// TwinCAT 3 PLC project Untitled1
// ProgramVersion: 3.1.4026.26
// project tree:
//   GVLs/HMI/ CNV_HMI.TcGVL, CNV_HMI_IO.TcGVL, GVL_HMI_Carousel.TcGVL, GVL_HMI_CNV.TcGVL, GVL_HMI_Gates.TcGVL, GVL_HMI_System.TcGVL, GVL_HMI_VTD.TcGVL
//   GVLs/IO/ IO_Cards.TcGVL, IO_Chargers.TcGVL, IO_RemoteModules.TcGVL, IO_Safety.TcGVL, IO_VFDs.TcGVL

// ---- GVLs/HMI/CNV_HMI.TcGVL
{attribute 'qualified_only'}
VAR_GLOBAL
	CNV_ID_HMI_Old_1:  DINT;
	CNV_ID_HMI:  DINT;
	CNV_ID_HMI_1:  DINT;
	CNV_ID_HMI_Old:  DInt;
	CNV_In_Out_1:  BOOL;
	CNV_Level_Selected:  UInt;
	CNV_Level_Selected_OLD:  UInt;
	CNV_Motor_Actual_Torque:  Real;
	CNV_Motor_Actual_Torque_1:  REAL;
	CNV_Motor_Current_Actual_HMI:  Real;
	CNV_Motor_Current_Actual_HMI_1:  REAL;
	CNV_Motor_Ready:  Bool;
	CNV_Motor_Ready_1:  BOOL;
	CNV_Motor_Status_HMI:  UInt;
	CNV_Motor_Status_HMI_1:  UINT;
	Cnv_Occupied_HMI:  Bool;
	Cnv_Occupied_HMI_1:  BOOL;
	CNV_System_Selected:  UInt;
	CVTD_CNV2_Selected:  UInt;
	Enable_HMI:  Bool;
	Enable_HMI_1:  Bool;
	Enabled_HMI:  Bool;
	Enabled_HMI_1:  Bool;
	Error_HMI:  Bool;
	Error_HMI_1:  Bool;
	HMI_Light_Guard_Bypass:  Bool;
	Light_Guard_Bypass_1:  Bool;
	Light_Guard_Bypass_2:  Bool;
	Manual_Bwd_HMI:  Bool;
	Manual_Bwd_HMI_1:  Bool;
	Manual_Fwd_HMI:  Bool;
	Manual_Fwd_HMI_1:  Bool;
	Manual_Sfty_Stopper_Down_1:  Bool;
	Manual_Sfty_Stopper_Up_1:  Bool;
	Mode_Change_HMI:  UInt;
	Mode_Change_HMI_1:  UInt;
	Mode_HMI:  UInt;
	Mode_HMI_1:  UInt;
	Motor_Direction_HMI:  UInt;
	Motor_Direction_HMI_1:  UInt;
	Motor_Speed_Actual_HMI:  UInt;
	Motor_Speed_Actual_HMI_1:  UInt;
	Motor_Speed_Requested_HMI:  UInt;
	Motor_Speed_Requested_HMI_1:  UInt;
	Ready_For_Task_HMI:  Bool;
	Ready_For_Task_HMI_1:  Bool;
	Reset_HMI:  Bool;
	Reset_HMI_1:  Bool;
	Running_HMI:  Bool;
	Running_HMI_1:  Bool;
	SM_State_HMI:  UInt;
	SM_State_HMI_1:  UInt;
	Start_Transfer_HMI:  Bool;
	Start_Transfer_HMI_1:  Bool;
	Stop_HMI:  Bool;
	Stopped_HMI:  Bool;
	Stopped_HMI_1:  Bool;
	Transfer_From_ID_HMI:  DInt;
	Transfer_From_ID_HMI_1:  DInt;
	Transfer_To_ID_HMI:  DInt;
	Transfer_To_ID_HMI_1:  DInt;
	UpDown_1:  UInt;
	Warning_HMI:  UInt;
	Warning_HMI_1:  UINT;
END_VAR

// ---- GVLs/HMI/CNV_HMI_IO.TcGVL
{attribute 'qualified_only'}
VAR_GLOBAL
	HMI_CNV_SftyPinDown_1:  BOOL;
	HMI_CNV_SftyPinUp_1:  BOOL;
	HMI_Light_Guard:  Bool;
	HMI_CNV_Forward_1:  Bool;
	HMI_CNV_Backward:  Bool;
	HMI_CNV_Forward:  Bool;
	HMI_CNV_Backward_1:  Bool;
END_VAR

// ---- GVLs/HMI/GVL_HMI_Carousel.TcGVL
// HMI interface of the screen Carrousel.
// Device index: 1..2 = PopUp 1..2, 3..7 = Roller 1..5, 8 = Chain, 9 = Turntable.
// TODO: FC_CarouselHmiUpdate once the carousel DUTs / FBs exist. Until then all values stay 0/FALSE.
{attribute 'qualified_only'}
VAR_GLOBAL
    uiSelected : UINT;                                   // HMI -> PLC: 1..9, see above
    astDevice : ARRAY[1..9] OF ST_HMI_ConveyorStatus;    // PLC -> HMI
    stSelected : ST_HMI_ConveyorStatus;                  // PLC -> HMI: copy of the selected device
    stCommand : ST_HMI_ConveyorCommand;                  // HMI -> PLC: commands for the selected device
END_VAR

// ---- GVLs/HMI/GVL_HMI_CNV.TcGVL
// HMI interface of the screen CNV (extractor + buffer conveyors L1..L6).
// The visualization uses only these variables.
// TODO: FC_CnvHmiUpdate (status from Control.ECnv / Control.LCnv, commands to the selected conveyor)
// once the Control refactor compiles. Until then all values stay 0/FALSE.
{attribute 'qualified_only'}
VAR_GLOBAL
    uiSelected : UINT;                                   // HMI -> PLC: 0 = extractor, 1..6 = buffer level
    astConveyor : ARRAY[0..6] OF ST_HMI_ConveyorStatus;  // PLC -> HMI: 0 = extractor, 1..6 = buffer L1..L6
    stSelected : ST_HMI_ConveyorStatus;                  // PLC -> HMI: copy of the selected conveyor
    stCommand : ST_HMI_ConveyorCommand;                  // HMI -> PLC: commands for the selected conveyor
END_VAR

// ---- GVLs/HMI/GVL_HMI_Gates.TcGVL
// HMI interface of the screen Access_Gates. Requests only; the gate locks are
// controlled by the safety logic (TwinSAFE / Euchner MGB2).
// TODO: FC_GatesHmiUpdate (status from Control.Gate_Station). Until then all values stay 0/FALSE.
{attribute 'qualified_only'}
VAR_GLOBAL
    astGate : ARRAY[1..2] OF ST_HMI_GateStatus;      // PLC -> HMI
    astCommand : ARRAY[1..2] OF ST_HMI_GateCommand;  // HMI -> PLC
END_VAR

// ---- GVLs/HMI/GVL_HMI_System.TcGVL
// HMI interface of the system overview (screen Main). The visualization uses only
// these variables; it must not access Control, IO GVLs or FB instances directly.
// TODO: FC_SystemHmiUpdateStatus fills the status from Control once the Control
// refactor (single VTD, carousel DUTs) compiles. Until then all values stay 0/FALSE.
{attribute 'qualified_only'}
VAR_GLOBAL
    stStatus : ST_HMI_SystemStatus;                    // PLC -> HMI
    stCommand : ST_HMI_SystemCommand;                  // HMI -> PLC
    stVtd : ST_HMI_VtdOverview;                        // PLC -> HMI
    stExtractor : ST_HMI_DeviceSummary;                // PLC -> HMI
    astBuffer : ARRAY[1..6] OF ST_HMI_DeviceSummary;   // PLC -> HMI, buffer levels L1..L6
    astPopUp : ARRAY[1..2] OF ST_HMI_DeviceSummary;    // PLC -> HMI, carousel popups
    astRoller : ARRAY[1..5] OF ST_HMI_DeviceSummary;   // PLC -> HMI, carousel rollers
    stChain : ST_HMI_DeviceSummary;                    // PLC -> HMI, carousel chain transfer
    stTurntable : ST_HMI_DeviceSummary;                // PLC -> HMI
    astGate : ARRAY[1..2] OF ST_HMI_GateSummary;       // PLC -> HMI
END_VAR

// ---- GVLs/HMI/GVL_HMI_VTD.TcGVL
// HMI interface of the VTD. The visualization uses only these variables;
// it must not access IO GVLs or FB instances directly.
{attribute 'qualified_only'}
VAR_GLOBAL
    // Screen "Visualization" - process data test (TEST ONLY)
    stPdStatus : ST_VTD_PdHmiStatus;   // PLC -> HMI, written by FC_VTD_PdHmiUpdateStatus
    stPdCommand : ST_VTD_PdHmiCommand; // HMI -> PLC, read by MAIN (TEST ONLY)

    // Screen "VTD_ManualTest" - manual control (TEST ONLY)
    stManualCommand : ST_VTD_ManualHmiCommand; // HMI -> PLC, read and partly written back by FB_VTD_ManualControl
    stManualStatus : ST_VTD_ManualHmiStatus;   // PLC -> HMI, written by MAIN

    // Screen "VTD" - operation
    stStatus : ST_HMI_VtdStatus;     // PLC -> HMI (TODO: FC_VtdHmiUpdate after the Control refactor)
    stCommand : ST_HMI_VtdCommand;   // HMI -> PLC
END_VAR

VAR_GLOBAL PERSISTENT
    stManualSettings : ST_VTD_ManualSettings;  // HMI <-> PLC, test settings kept over a restart
END_VAR

// ---- GVLs/IO/IO_Cards.TcGVL
{attribute 'qualified_only'}
VAR_GLOBAL
	// Source: INBOUND VTD ELECTRICAL DRAWING_9_17_26.pdf, sheets 24.0-27.0.
	// Local PLC rack cards only. Remote module signals belong in a separate IO_Remote GVL.
	// Channel comments identify physical terminals, not PLC process-image offsets.
	// AT %I* / AT %Q* declarations require individual channel links in TwinCAT XAE.
	// Spare outputs are reserved; do not use them in control logic.

	// DI-01 (EL1809) - card 23.0-1, sheet 24.0.
	// Existing REDUNDANCY_OK_8PS1 name retained; the drawing identifies redundancy module 8RS1.
	REDUNDANCY_OK_8PS1 AT %I* : BOOL; // DI-01 CH01 | Wire 24.01 | 8RS1 redundancy OK
	HANDHELD_HMI_KEY_SWITCH_1_NO AT %I* : BOOL; // DI-01 CH02 | Wire 24.02
	HANDHELD_HMI_KEY_SWITCH_2_NO AT %I* : BOOL; // DI-01 CH03 | Wire 24.03
	HANDHELD_HMI_CONNECTED AT %I* : BOOL; // DI-01 CH04 | Wire 24.04
	LM3_4_FAULT AT %I* : BOOL; // DI-01 CH05 | Wire 24.05
	LM5_6_FAULT AT %I* : BOOL; // DI-01 CH06 | Wire 24.06
	LM7_8_FAULT AT %I* : BOOL; // DI-01 CH07 | Wire 24.07
	LM9_FAULT AT %I* : BOOL; // DI-01 CH08 | Wire 24.08
	LM10_FAULT AT %I* : BOOL; // DI-01 CH09 | Wire 24.09
	LM11_FAULT AT %I* : BOOL; // DI-01 CH10 | Wire 24.10
	LM12_FAULT AT %I* : BOOL; // DI-01 CH11 | Wire 24.11
	LM13_14_FAULT AT %I* : BOOL; // DI-01 CH12 | Wire 24.12
	LM15_FAULT AT %I* : BOOL; // DI-01 CH13 | Wire 24.13
	
	LM16_FAULT AT %I* : BOOL; // DI-01 CH14 | Wire 24.14
	_8PS1_OUT_100 AT %I* : BOOL; // DI-01 CH15 | Wire 24.15
	_8PS1_DC_OK AT %I* : BOOL; // DI-01 CH16 | Wire 24.16

	// DI-02 (EL1809) - card 23.0-2, sheet 25.0.
	BACKUP_SIGNAL_BU AT %I* : BOOL; // DI-02 CH01 | Wire 25.01
	TROUBLE_SIGNAL_TR AT %I* : BOOL; // DI-02 CH02 | Wire 25.02
	BATTERY_LOW_SIGNAL_BL AT %I* : BOOL; // DI-02 CH03 | Wire 25.03
	BATTERY_REPLACEMENT_WB AT %I* : BOOL; // DI-02 CH04 | Wire 25.04
	_8PS2_100 AT %I* : BOOL; // DI-02 CH05 | Wire 25.05
	_8PS2_DC_OK AT %I* : BOOL; // DI-02 CH06 | Wire 25.06
	_8PS3_100 AT %I* : BOOL; // DI-02 CH07 | Wire 25.07
	_8PS3_DC_OK AT %I* : BOOL; // DI-02 CH08 | Wire 25.08
	LM100_FAULT AT %I* : BOOL; // DI-02 CH09 | Wire 25.09
	LM101_FAULT AT %I* : BOOL; // DI-02 CH10 | Wire 25.10
	LM102_FAULT AT %I* : BOOL; // DI-02 CH11 | Wire 25.11
	LM103_FAULT AT %I* : BOOL; // DI-02 CH12 | Wire 25.12
	LM104_FAULT AT %I* : BOOL; // DI-02 CH13 | Wire 25.13
	LM105_FAULT AT %I* : BOOL; // DI-02 CH14 | Wire 25.14
	LM106_FAULT AT %I* : BOOL; // DI-02 CH15 | Wire 25.15
	LM107_FAULT AT %I* : BOOL; // DI-02 CH16 | Wire 25.16

	// DO-01 (EL2809) - card 23.0-3, sheet 26.0.
	LM3_16_SET_RESET AT %Q* : BOOL; // DO-01 CH01 | Wire 26.01 | Relay 26CR1
	_50K50_BEACON_INDICATOR_RED AT %Q* : BOOL; // DO-01 CH02 | Wire 26.02 | Relay 26CR2
	_50K50_BEACON_INDICATOR_YELLOW AT %Q* : BOOL; // DO-01 CH03 | Wire 26.03 | Relay 26CR3
	_50K50_BEACON_INDICATOR_GREEN AT %Q* : BOOL; // DO-01 CH04 | Wire 26.04 | Relay 26CR4
	_50K50_BEACON_BUZZER AT %Q* : BOOL; // DO-01 CH05 | Wire 26.05 | Relay 26CR5
	LM100_107_SET_RESET AT %Q* : BOOL; // DO-01 CH06 | Wire 26.06 | Relay 26CR6
	BYPASS_1_FROM_DIGITAL_PLC_OUTPUT AT %Q* : BOOL; // DO-01 CH07 | Wire 26.07 | Relay 26CR7 | Existing safety-interface signal; no bypass logic added
	BYPASS_2_FROM_DIGITAL_PLC_OUTPUT AT %Q* : BOOL; // DO-01 CH08 | Wire 26.08 | Relay 26CR8 | Existing safety-interface signal; no bypass logic added
	BUZZER AT %Q* : BOOL; // DO-01 CH09 | Wire 26.09 | Relay 26CR9
	DO_01_SPARE_CH10 AT %Q* : BOOL; // DO-01 CH10 | Wire 26.10 | Relay 26CR10 | Spare
	DO_01_SPARE_CH11 AT %Q* : BOOL; // DO-01 CH11 | Wire 26.11 | Relay 26CR11 | Spare
	DO_01_SPARE_CH12 AT %Q* : BOOL; // DO-01 CH12 | Wire 26.12 | Relay 26CR12 | Spare
	DO_01_SPARE_CH13 AT %Q* : BOOL; // DO-01 CH13 | Wire 26.13 | Relay 26CR13 | Spare
	DO_01_SPARE_CH14 AT %Q* : BOOL; // DO-01 CH14 | Wire 26.14 | Relay 26CR14 | Spare
	DO_01_SPARE_CH15 AT %Q* : BOOL; // DO-01 CH15 | Wire 26.15 | Relay 26CR15 | Spare
	DO_01_SPARE_CH16 AT %Q* : BOOL; // DO-01 CH16 | Wire 26.16 | Relay 26CR16 | Spare

	// DO-02 (EL2809) - card 23.0-4, sheet 27.0.
	// UPS control uses CH15/CH16. CH01-CH14 are spare.
	DO_02_SPARE_CH01 AT %Q* : BOOL; // DO-02 CH01 | Wire 27.01 | Relay 27CR1 | Spare
	DO_02_SPARE_CH02 AT %Q* : BOOL; // DO-02 CH02 | Wire 27.02 | Relay 27CR2 | Spare
	DO_02_SPARE_CH03 AT %Q* : BOOL; // DO-02 CH03 | Wire 27.03 | Relay 27CR3 | Spare
	DO_02_SPARE_CH04 AT %Q* : BOOL; // DO-02 CH04 | Wire 27.04 | Relay 27CR4 | Spare
	DO_02_SPARE_CH05 AT %Q* : BOOL; // DO-02 CH05 | Wire 27.05 | Relay 27CR5 | Spare
	DO_02_SPARE_CH06 AT %Q* : BOOL; // DO-02 CH06 | Wire 27.06 | Relay 27CR6 | Spare
	DO_02_SPARE_CH07 AT %Q* : BOOL; // DO-02 CH07 | Wire 27.07 | Relay 27CR7 | Spare
	DO_02_SPARE_CH08 AT %Q* : BOOL; // DO-02 CH08 | Wire 27.08 | Relay 27CR8 | Spare
	DO_02_SPARE_CH09 AT %Q* : BOOL; // DO-02 CH09 | Wire 27.09 | Relay 27CR9 | Spare
	DO_02_SPARE_CH10 AT %Q* : BOOL; // DO-02 CH10 | Drawing labels wire 27.27 and relay 27CR27; verify drawing tag. | Spare
	DO_02_SPARE_CH11 AT %Q* : BOOL; // DO-02 CH11 | Wire 27.11 | Relay 27CR11 | Spare
	DO_02_SPARE_CH12 AT %Q* : BOOL; // DO-02 CH12 | Wire 27.12 | Relay 27CR12 | Spare
	DO_02_SPARE_CH13 AT %Q* : BOOL; // DO-02 CH13 | Wire 27.13 | Relay 27CR13 | Spare
	DO_02_SPARE_CH14 AT %Q* : BOOL; // DO-02 CH14 | Wire 27.14 | Relay 27CR14 | Spare
	_8BPS1_REMOTE_ON_OFF AT %Q* : BOOL; // DO-02 CH15 | Wire 27.15 | Relay 27CR15
	_8BPS1_BACKUP_STOP AT %Q* : BOOL; // DO-02 CH16 | Wire 27.16 | Relay 27CR16

	// Existing safety-related declarations below are preserved for compatibility.
	// These standard PLC BOOLs do not implement a safety function.
	// Their relationship to validated TwinSAFE diagnostics must be reviewed before use.
	// See docs/IO_Cards_Review.md for the complete EL1918/EL2912 drawing inventory.
	//FDI-01 (EL1918) - SAFETY INPUTS 23.0-6
	EMERGENCY_STOP_ON_DOOR_CH1 AT%I*:BOOL;
	EMERGENCY_STOP_ON_DOOR_CH2 AT%I*:BOOL;
	EMERGENCY_STOP_ON_HMI AT%I*:BOOL;
END_VAR

// ---- GVLs/IO/IO_Chargers.TcGVL
{attribute 'qualified_only'}
VAR_GLOBAL
// 	Charger Level 1
	Inputs_1 AT%I*:ARRAY[0..19] OF BYTE;
	Outputs_1 AT%Q*:ARRAY[0..9] OF BYTE;
	
	// 	Charger Level 2
	Inputs_2 AT%I*:ARRAY[0..19] OF BYTE;
	Outputs_2 AT%Q*:ARRAY[0..9] OF BYTE;
	
	// 	Charger Level 3
	Inputs_3 AT%I*:ARRAY[0..19] OF BYTE;
	Outputs_3 AT%Q*:ARRAY[0..9] OF BYTE;
	
	// 	Charger Level 4
	Inputs_4 AT%I*:ARRAY[0..19] OF BYTE;
	Outputs_4 AT%Q*:ARRAY[0..9] OF BYTE;
	
	// 	Charger Level 5
	Inputs_5 AT%I*:ARRAY[0..19] OF BYTE;
	Outputs_5 AT%Q*:ARRAY[0..9] OF BYTE;
	
	// 	Charger Level 6
	Inputs_6 AT%I*:ARRAY[0..19] OF BYTE;
	Outputs_6 AT%Q*:ARRAY[0..9] OF BYTE;
	
	// 	Charger Level 7
	Inputs_7 AT%I*:ARRAY[0..19] OF BYTE;
	Outputs_7 AT%Q*:ARRAY[0..9] OF BYTE;
	
	// 	Charger Level 8
	Inputs_8 AT%I*:ARRAY[0..19] OF BYTE;
	Outputs_8 AT%Q*:ARRAY[0..9] OF BYTE;	
END_VAR

// ---- GVLs/IO/IO_RemoteModules.TcGVL
{attribute 'qualified_only'}
VAR_GLOBAL
    // Source: INBOUND VTD ELECTRICAL DRAWING_9_17_26.pdf (rev D), sheets 43.0-48.6 and 53.0-53.5.
    // EtherCAT P remote I/O boxes and TwinSAFE boxes. Local rack cards are in IO_Cards.
    // Box headers give the TwinCAT box name (SpaceX.tsproj) and the drawing tag. The box-to-tag
    // mapping follows the numbering order (confirmed by the user, 2026-10-21).
    // Channel comments: <drawing tag> CH<nn> | <connector> | <description>.
    //   EPP1008: one input per M12 socket X01-X08 (pin 4).
    //   EPP1809: two inputs per M12 socket, X01-X16 (first channel pin 4, second channel pin 2).
    //   EPP2328: four M12 sockets; channel A = pin 4, channel B = pin 2 (sheet 53.0 pinout).
    // AT %I* / AT %Q* declarations require individual channel links in TwinCAT XAE.
    // Spare and unnamed channels are reserved; do not use them in control logic.
    // EtherCAT diagnostics (WcState / EcState) are not linked yet: link them manually in XAE.

    // ---------------------------------------------------------------- Carousel conveyors, EPP1008-0022
    // Sheets 45.0-45.1 / 46.0: boxes for carousel conveyor popups 1-2 and turntable + roller.
    // All EPP1008 channels are shown as '?????????' in drawing rev D: declared as reserved,
    // rename them when the drawing names the signals.
    // 45RIO4 = ENCODER (EPP5001-0002), turntable SSI encoder, sheet 45.5: not part of this GVL.

    // DI-01 (EPP1008-0022) = 45RIO1 - carousel conveyors area section 3 - sheet 45.2.
    _45RIO1_CH01 AT %I* : BOOL; // 45RIO1 CH01 | X01 | Not named in drawing rev D
    _45RIO1_CH02 AT %I* : BOOL; // 45RIO1 CH02 | X02 | Not named in drawing rev D
    _45RIO1_CH03 AT %I* : BOOL; // 45RIO1 CH03 | X03 | Not named in drawing rev D
    _45RIO1_CH04 AT %I* : BOOL; // 45RIO1 CH04 | X04 | Not named in drawing rev D
    _45RIO1_CH05 AT %I* : BOOL; // 45RIO1 CH05 | X05 | Not named in drawing rev D
    _45RIO1_CH06 AT %I* : BOOL; // 45RIO1 CH06 | X06 | Not named in drawing rev D
    _45RIO1_CH07 AT %I* : BOOL; // 45RIO1 CH07 | X07 | Not named in drawing rev D
    _45RIO1_CH08 AT %I* : BOOL; // 45RIO1 CH08 | X08 | Not named in drawing rev D
    _45RIO1_WcState AT %I* : BOOL; // DI-01 > WcState > WcState (TRUE = data invalid)
    _45RIO1_EcState AT %I* : UINT; // DI-01 > InfoData > State (8 = OP)

    // DI-02 (EPP1008-0022) = 45RIO2 - carousel conveyors area section 3 - sheet 45.3.
    _45RIO2_CH01 AT %I* : BOOL; // 45RIO2 CH01 | X01 | Not named in drawing rev D
    _45RIO2_CH02 AT %I* : BOOL; // 45RIO2 CH02 | X02 | Not named in drawing rev D
    _45RIO2_CH03 AT %I* : BOOL; // 45RIO2 CH03 | X03 | Not named in drawing rev D
    _45RIO2_CH04 AT %I* : BOOL; // 45RIO2 CH04 | X04 | Not named in drawing rev D
    _45RIO2_CH05 AT %I* : BOOL; // 45RIO2 CH05 | X05 | Not named in drawing rev D
    _45RIO2_CH06 AT %I* : BOOL; // 45RIO2 CH06 | X06 | Not named in drawing rev D
    _45RIO2_CH07 AT %I* : BOOL; // 45RIO2 CH07 | X07 | Not named in drawing rev D
    _45RIO2_CH08 AT %I* : BOOL; // 45RIO2 CH08 | X08 | Not named in drawing rev D
    _45RIO2_WcState AT %I* : BOOL; // DI-02 > WcState > WcState (TRUE = data invalid)
    _45RIO2_EcState AT %I* : UINT; // DI-02 > InfoData > State (8 = OP)

    // DI-03 (EPP1008-0022) = 45RIO3 - carousel conveyors area section 3 - sheet 45.4.
    _45RIO3_CH01 AT %I* : BOOL; // 45RIO3 CH01 | X01 | Not named in drawing rev D
    _45RIO3_CH02 AT %I* : BOOL; // 45RIO3 CH02 | X02 | Not named in drawing rev D
    _45RIO3_CH03 AT %I* : BOOL; // 45RIO3 CH03 | X03 | Not named in drawing rev D
    _45RIO3_CH04 AT %I* : BOOL; // 45RIO3 CH04 | X04 | Not named in drawing rev D
    _45RIO3_CH05 AT %I* : BOOL; // 45RIO3 CH05 | X05 | Not named in drawing rev D
    _45RIO3_CH06 AT %I* : BOOL; // 45RIO3 CH06 | X06 | Not named in drawing rev D
    _45RIO3_CH07 AT %I* : BOOL; // 45RIO3 CH07 | X07 | Not named in drawing rev D
    _45RIO3_CH08 AT %I* : BOOL; // 45RIO3 CH08 | X08 | Not named in drawing rev D
    _45RIO3_WcState AT %I* : BOOL; // DI-03 > WcState > WcState (TRUE = data invalid)
    _45RIO3_EcState AT %I* : UINT; // DI-03 > InfoData > State (8 = OP)

    // DI-04 (EPP1008-0022) = 46RIO1 - carousel conveyors area sections 1 & 2 - sheet 46.1.
    _46RIO1_CH01 AT %I* : BOOL; // 46RIO1 CH01 | X01 | Not named in drawing rev D
    _46RIO1_CH02 AT %I* : BOOL; // 46RIO1 CH02 | X02 | Not named in drawing rev D
    _46RIO1_CH03 AT %I* : BOOL; // 46RIO1 CH03 | X03 | Not named in drawing rev D
    _46RIO1_CH04 AT %I* : BOOL; // 46RIO1 CH04 | X04 | Not named in drawing rev D
    _46RIO1_CH05 AT %I* : BOOL; // 46RIO1 CH05 | X05 | Not named in drawing rev D
    _46RIO1_CH06 AT %I* : BOOL; // 46RIO1 CH06 | X06 | Not named in drawing rev D
    _46RIO1_CH07 AT %I* : BOOL; // 46RIO1 CH07 | X07 | Not named in drawing rev D
    _46RIO1_CH08 AT %I* : BOOL; // 46RIO1 CH08 | X08 | Not named in drawing rev D
    _46RIO1_WcState AT %I* : BOOL; // DI-04 > WcState > WcState (TRUE = data invalid)
    _46RIO1_EcState AT %I* : UINT; // DI-04 > InfoData > State (8 = OP)

    // DI-05 (EPP1008-0022) = 46RIO2 - carousel conveyors area sections 1 & 2 - sheet 46.2.
    _46RIO2_CH01 AT %I* : BOOL; // 46RIO2 CH01 | X01 | Not named in drawing rev D
    _46RIO2_CH02 AT %I* : BOOL; // 46RIO2 CH02 | X02 | Not named in drawing rev D
    _46RIO2_CH03 AT %I* : BOOL; // 46RIO2 CH03 | X03 | Not named in drawing rev D
    _46RIO2_CH04 AT %I* : BOOL; // 46RIO2 CH04 | X04 | Not named in drawing rev D
    _46RIO2_CH05 AT %I* : BOOL; // 46RIO2 CH05 | X05 | Not named in drawing rev D
    _46RIO2_CH06 AT %I* : BOOL; // 46RIO2 CH06 | X06 | Not named in drawing rev D
    _46RIO2_CH07 AT %I* : BOOL; // 46RIO2 CH07 | X07 | Not named in drawing rev D
    _46RIO2_CH08 AT %I* : BOOL; // 46RIO2 CH08 | X08 | Not named in drawing rev D
    _46RIO2_WcState AT %I* : BOOL; // DI-05 > WcState > WcState (TRUE = data invalid)
    _46RIO2_EcState AT %I* : UINT; // DI-05 > InfoData > State (8 = OP)

    // DI-06 (EPP1008-0022) = 46RIO3 - carousel conveyors area sections 1 & 2 - sheet 46.3.
    _46RIO3_CH01 AT %I* : BOOL; // 46RIO3 CH01 | X01 | Not named in drawing rev D
    _46RIO3_CH02 AT %I* : BOOL; // 46RIO3 CH02 | X02 | Not named in drawing rev D
    _46RIO3_CH03 AT %I* : BOOL; // 46RIO3 CH03 | X03 | Not named in drawing rev D
    _46RIO3_CH04 AT %I* : BOOL; // 46RIO3 CH04 | X04 | Not named in drawing rev D
    _46RIO3_CH05 AT %I* : BOOL; // 46RIO3 CH05 | X05 | Not named in drawing rev D
    _46RIO3_CH06 AT %I* : BOOL; // 46RIO3 CH06 | X06 | Not named in drawing rev D
    _46RIO3_CH07 AT %I* : BOOL; // 46RIO3 CH07 | X07 | Not named in drawing rev D
    _46RIO3_CH08 AT %I* : BOOL; // 46RIO3 CH08 | X08 | Not named in drawing rev D
    _46RIO3_WcState AT %I* : BOOL; // DI-06 > WcState > WcState (TRUE = data invalid)
    _46RIO3_EcState AT %I* : UINT; // DI-06 > InfoData > State (8 = OP)

    // DI-07 (EPP1008-0022) = 46RIO4 - carousel conveyors area sections 1 & 2 - sheet 46.4.
    _46RIO4_CH01 AT %I* : BOOL; // 46RIO4 CH01 | X01 | Not named in drawing rev D
    _46RIO4_CH02 AT %I* : BOOL; // 46RIO4 CH02 | X02 | Not named in drawing rev D
    _46RIO4_CH03 AT %I* : BOOL; // 46RIO4 CH03 | X03 | Not named in drawing rev D
    _46RIO4_CH04 AT %I* : BOOL; // 46RIO4 CH04 | X04 | Not named in drawing rev D
    _46RIO4_CH05 AT %I* : BOOL; // 46RIO4 CH05 | X05 | Not named in drawing rev D
    _46RIO4_CH06 AT %I* : BOOL; // 46RIO4 CH06 | X06 | Not named in drawing rev D
    _46RIO4_CH07 AT %I* : BOOL; // 46RIO4 CH07 | X07 | Not named in drawing rev D
    _46RIO4_CH08 AT %I* : BOOL; // 46RIO4 CH08 | X08 | Not named in drawing rev D
    _46RIO4_WcState AT %I* : BOOL; // DI-07 > WcState > WcState (TRUE = data invalid)
    _46RIO4_EcState AT %I* : UINT; // DI-07 > InfoData > State (8 = OP)

    // DI-08 (EPP1008-0022) = 46RIO5 - carousel conveyors area sections 1 & 2 - sheet 46.5.
    _46RIO5_CH01 AT %I* : BOOL; // 46RIO5 CH01 | X01 | Not named in drawing rev D
    _46RIO5_CH02 AT %I* : BOOL; // 46RIO5 CH02 | X02 | Not named in drawing rev D
    _46RIO5_CH03 AT %I* : BOOL; // 46RIO5 CH03 | X03 | Not named in drawing rev D
    _46RIO5_CH04 AT %I* : BOOL; // 46RIO5 CH04 | X04 | Not named in drawing rev D
    _46RIO5_CH05 AT %I* : BOOL; // 46RIO5 CH05 | X05 | Not named in drawing rev D
    _46RIO5_CH06 AT %I* : BOOL; // 46RIO5 CH06 | X06 | Not named in drawing rev D
    _46RIO5_CH07 AT %I* : BOOL; // 46RIO5 CH07 | X07 | Not named in drawing rev D
    _46RIO5_CH08 AT %I* : BOOL; // 46RIO5 CH08 | X08 | Not named in drawing rev D
    _46RIO5_WcState AT %I* : BOOL; // DI-08 > WcState > WcState (TRUE = data invalid)
    _46RIO5_EcState AT %I* : UINT; // DI-08 > InfoData > State (8 = OP)

    // DI-09 (EPP1008-0022) = 46RIO6 - carousel conveyors area sections 1 & 2 - sheet 46.6.
    _46RIO6_CH01 AT %I* : BOOL; // 46RIO6 CH01 | X01 | Not named in drawing rev D
    _46RIO6_CH02 AT %I* : BOOL; // 46RIO6 CH02 | X02 | Not named in drawing rev D
    _46RIO6_CH03 AT %I* : BOOL; // 46RIO6 CH03 | X03 | Not named in drawing rev D
    _46RIO6_CH04 AT %I* : BOOL; // 46RIO6 CH04 | X04 | Not named in drawing rev D
    _46RIO6_CH05 AT %I* : BOOL; // 46RIO6 CH05 | X05 | Not named in drawing rev D
    _46RIO6_CH06 AT %I* : BOOL; // 46RIO6 CH06 | X06 | Not named in drawing rev D
    _46RIO6_CH07 AT %I* : BOOL; // 46RIO6 CH07 | X07 | Not named in drawing rev D
    _46RIO6_CH08 AT %I* : BOOL; // 46RIO6 CH08 | X08 | Not named in drawing rev D
    _46RIO6_WcState AT %I* : BOOL; // DI-09 > WcState > WcState (TRUE = data invalid)
    _46RIO6_EcState AT %I* : UINT; // DI-09 > InfoData > State (8 = OP)

    // DI-10 (EPP1008-0022) = 46RIO7 - carousel conveyors area sections 1 & 2 - sheet 46.7.
    _46RIO7_CH01 AT %I* : BOOL; // 46RIO7 CH01 | X01 | Not named in drawing rev D
    _46RIO7_CH02 AT %I* : BOOL; // 46RIO7 CH02 | X02 | Not named in drawing rev D
    _46RIO7_CH03 AT %I* : BOOL; // 46RIO7 CH03 | X03 | Not named in drawing rev D
    _46RIO7_CH04 AT %I* : BOOL; // 46RIO7 CH04 | X04 | Not named in drawing rev D
    _46RIO7_CH05 AT %I* : BOOL; // 46RIO7 CH05 | X05 | Not named in drawing rev D
    _46RIO7_CH06 AT %I* : BOOL; // 46RIO7 CH06 | X06 | Not named in drawing rev D
    _46RIO7_CH07 AT %I* : BOOL; // 46RIO7 CH07 | X07 | Not named in drawing rev D
    _46RIO7_CH08 AT %I* : BOOL; // 46RIO7 CH08 | X08 | Not named in drawing rev D
    _46RIO7_WcState AT %I* : BOOL; // DI-10 > WcState > WcState (TRUE = data invalid)
    _46RIO7_EcState AT %I* : UINT; // DI-10 > InfoData > State (8 = OP)

    // ---------------------------------------------------------------- Docking pins and VTD detection

    // DIO-01 (EPP2328-0002) = 47RIO1 - docking pins - sheet 47.3.
    // Outputs go to the docking pins junction box (separate drawing, see note on sheet 47.3).
    // Two signals per socket through Y-cables 6ES7194-6KA00-0XA0 (legs II / III):
    // confirm the leg-to-channel order at the I/O check.
    LEFT_LOCKING_PINS_EXTENDED AT %I* : BOOL; // 47RIO1 CH01 | M12-1 pin 4 | From left locking pins extended proximity sensors
    RIGHT_LOCKING_PINS_EXTENDED AT %I* : BOOL; // 47RIO1 CH02 | M12-1 pin 2 | From right locking pins extended proximity sensors
    LEFT_LOCKING_PINS_RETRACTED AT %I* : BOOL; // 47RIO1 CH03 | M12-2 pin 4 | From left locking pins retracted proximity sensors
    RIGHT_LOCKING_PINS_RETRACTED AT %I* : BOOL; // 47RIO1 CH04 | M12-2 pin 2 | From right locking pins retracted proximity sensors
    DOCKING_PINS_3KA1 AT %Q* : BOOL; // 47RIO1 CH05 | M12-3 pin 4 | To 3KA1 in docking pins junction box
    DOCKING_PINS_3KA2 AT %Q* : BOOL; // 47RIO1 CH06 | M12-3 pin 2 | To 3KA2 in docking pins junction box
    DOCKING_PINS_3KA3 AT %Q* : BOOL; // 47RIO1 CH07 | M12-4 pin 4 | To 3KA3 in docking pins junction box
    DOCKING_PINS_3KA4 AT %Q* : BOOL; // 47RIO1 CH08 | M12-4 pin 2 | To 3KA4 in docking pins junction box
    _47RIO1_WcState AT %I* : BOOL; // DIO-01 > WcState > WcState (TRUE = data invalid)
    _47RIO1_EcState AT %I* : UINT; // DIO-01 > InfoData > State (8 = OP)

    // DI-11 (EPP1809-0022) = 47RIO2 - VTD level, speed and pallet / shuttle detection - sheet 47.4.
    LEVEL_DETECT_1_SENSOR AT %I* : BOOL; // 47RIO2 CH01 | X01 | Level detect 1 sensor
    LEVEL_DETECT_2_SENSOR AT %I* : BOOL; // 47RIO2 CH02 | X02 | Level detect 2 sensor
    CREEP_SENSOR AT %I* : BOOL; // 47RIO2 CH03 | X03 | Creep sensor
    SLOWDOWN_SENSOR AT %I* : BOOL; // 47RIO2 CH04 | X04 | Slowdown sensor
    _47RIO2_CH05 AT %I* : BOOL; // 47RIO2 CH05 | X05 | Wired, not named in drawing rev D
    _47RIO2_SPARE_CH06 AT %I* : BOOL; // 47RIO2 CH06 | X06 | Spare
    _47RIO2_CH07 AT %I* : BOOL; // 47RIO2 CH07 | X07 | Wired, not named in drawing rev D
    _47RIO2_SPARE_CH08 AT %I* : BOOL; // 47RIO2 CH08 | X08 | Spare
    PALLET_DETECTION_1 AT %I* : BOOL; // 47RIO2 CH09 | X09 | Pallet detection #1
    PALLET_DETECTION_2 AT %I* : BOOL; // 47RIO2 CH10 | X10 | Pallet detection #2
    PALLET_DETECTION_3 AT %I* : BOOL; // 47RIO2 CH11 | X11 | Pallet detection #3
    PALLET_DETECTION_4 AT %I* : BOOL; // 47RIO2 CH12 | X12 | Pallet detection #4
    PALLET_DETECTION_5 AT %I* : BOOL; // 47RIO2 CH13 | X13 | Pallet detection #5
    PALLET_DETECTION_6 AT %I* : BOOL; // 47RIO2 CH14 | X14 | Pallet detection #6
    SHUTTLE_DETECTION_1 AT %I* : BOOL; // 47RIO2 CH15 | X15 | Shuttle detection #1
    SHUTTLE_DETECTION_2 AT %I* : BOOL; // 47RIO2 CH16 | X16 | Shuttle detection #2
    _47RIO2_WcState AT %I* : BOOL; // DI-11 > WcState > WcState (TRUE = data invalid)
    _47RIO2_EcState AT %I* : UINT; // DI-11 > InfoData > State (8 = OP)

    // ---------------------------------------------------------------- Buffer conveyors with stopper, EPP2328-0002
    // Outputs drive the coil of stopper motor relays SR8-BB-06A1 (sheets 53.0-53.5).

    // DIO-02 (EPP2328-0002) = 48RIO1 - conveyor with stopper, level 1 - sheets 48.1 and 53.0.
    BUFFER_L1_SAFETY_STOPPER_UPPER_SENSOR AT %I* : BOOL; // 48RIO1 CH01 | M12-1 pin 4 | Safety stopper upper sensor
    BUFFER_L1_SAFETY_STOPPER_LOWER_SENSOR AT %I* : BOOL; // 48RIO1 CH02 | M12-1 pin 2 | Safety stopper lower sensor
    BUFFER_L1_CONVEYOR_SENSOR_1 AT %I* : BOOL; // 48RIO1 CH03 | M12-2 pin 4 | Buffer conveyor sensor 1
    BUFFER_L1_CONVEYOR_SENSOR_2 AT %I* : BOOL; // 48RIO1 CH04 | M12-2 pin 2 | Buffer conveyor sensor 2
    BUFFER_L1_STOPPER_RELAY_53RR1 AT %Q* : BOOL; // 48RIO1 CH05 | M12-3 pin 4 | 53RR1 coil, stopper motor #1 53M1, sheet 53.0/5A
    _48RIO1_SPARE_CH06 AT %Q* : BOOL; // 48RIO1 CH06 | M12-3 pin 2 | Spare
    BUFFER_L1_STOPPER_RELAY_53RR2 AT %Q* : BOOL; // 48RIO1 CH07 | M12-4 pin 4 | 53RR2 coil, sheet 53.0/7E (relay not detailed in drawing rev D)
    _48RIO1_SPARE_CH08 AT %Q* : BOOL; // 48RIO1 CH08 | M12-4 pin 2 | Spare
    _48RIO1_WcState AT %I* : BOOL; // DIO-02 > WcState > WcState (TRUE = data invalid)
    _48RIO1_EcState AT %I* : UINT; // DIO-02 > InfoData > State (8 = OP)

    // DIO-03 (EPP2328-0002) = 48RIO2 - conveyor with stopper, level 2 - sheets 48.2 and 53.1.
    BUFFER_L2_SAFETY_STOPPER_UPPER_SENSOR AT %I* : BOOL; // 48RIO2 CH01 | M12-1 pin 4 | Safety stopper upper sensor
    BUFFER_L2_SAFETY_STOPPER_LOWER_SENSOR AT %I* : BOOL; // 48RIO2 CH02 | M12-1 pin 2 | Safety stopper lower sensor
    BUFFER_L2_CONVEYOR_SENSOR_1 AT %I* : BOOL; // 48RIO2 CH03 | M12-2 pin 4 | Buffer conveyor sensor 1
    BUFFER_L2_CONVEYOR_SENSOR_2 AT %I* : BOOL; // 48RIO2 CH04 | M12-2 pin 2 | Buffer conveyor sensor 2
    BUFFER_L2_STOPPER_RELAY_53RR3 AT %Q* : BOOL; // 48RIO2 CH05 | M12-3 pin 4 | 53RR3 coil, stopper motor #3 53M3, sheet 53.1/5A
    _48RIO2_SPARE_CH06 AT %Q* : BOOL; // 48RIO2 CH06 | M12-3 pin 2 | Spare
    BUFFER_L2_STOPPER_RELAY_53RR4 AT %Q* : BOOL; // 48RIO2 CH07 | M12-4 pin 4 | 53RR4 coil, sheet 53.1/7E (relay not detailed in drawing rev D)
    _48RIO2_SPARE_CH08 AT %Q* : BOOL; // 48RIO2 CH08 | M12-4 pin 2 | Spare
    _48RIO2_WcState AT %I* : BOOL; // DIO-03 > WcState > WcState (TRUE = data invalid)
    _48RIO2_EcState AT %I* : UINT; // DIO-03 > InfoData > State (8 = OP)

    // DIO-04 (EPP2328-0002) = 48RIO3 - conveyor with stopper, level 3 - sheets 48.3 and 53.2.
    BUFFER_L3_SAFETY_STOPPER_UPPER_SENSOR AT %I* : BOOL; // 48RIO3 CH01 | M12-1 pin 4 | Safety stopper upper sensor
    BUFFER_L3_SAFETY_STOPPER_LOWER_SENSOR AT %I* : BOOL; // 48RIO3 CH02 | M12-1 pin 2 | Safety stopper lower sensor
    BUFFER_L3_CONVEYOR_SENSOR_1 AT %I* : BOOL; // 48RIO3 CH03 | M12-2 pin 4 | Buffer conveyor sensor 1
    BUFFER_L3_CONVEYOR_SENSOR_2 AT %I* : BOOL; // 48RIO3 CH04 | M12-2 pin 2 | Buffer conveyor sensor 2
    BUFFER_L3_STOPPER_RELAY_53RR5 AT %Q* : BOOL; // 48RIO3 CH05 | M12-3 pin 4 | 53RR5 coil, stopper motor #5 53M5, sheet 53.2/5A
    _48RIO3_SPARE_CH06 AT %Q* : BOOL; // 48RIO3 CH06 | M12-3 pin 2 | Spare
    BUFFER_L3_STOPPER_RELAY_53RR6 AT %Q* : BOOL; // 48RIO3 CH07 | M12-4 pin 4 | 53RR6 coil, sheet 53.2/7E (relay not detailed in drawing rev D)
    _48RIO3_SPARE_CH08 AT %Q* : BOOL; // 48RIO3 CH08 | M12-4 pin 2 | Spare
    _48RIO3_WcState AT %I* : BOOL; // DIO-04 > WcState > WcState (TRUE = data invalid)
    _48RIO3_EcState AT %I* : UINT; // DIO-04 > InfoData > State (8 = OP)

    // DIO-05 (EPP2328-0002) = 48RIO4 - conveyor with stopper, level 4 - sheets 48.4 and 53.3.
    BUFFER_L4_SAFETY_STOPPER_UPPER_SENSOR AT %I* : BOOL; // 48RIO4 CH01 | M12-1 pin 4 | Safety stopper upper sensor
    BUFFER_L4_SAFETY_STOPPER_LOWER_SENSOR AT %I* : BOOL; // 48RIO4 CH02 | M12-1 pin 2 | Safety stopper lower sensor
    BUFFER_L4_CONVEYOR_SENSOR_1 AT %I* : BOOL; // 48RIO4 CH03 | M12-2 pin 4 | Buffer conveyor sensor 1
    BUFFER_L4_CONVEYOR_SENSOR_2 AT %I* : BOOL; // 48RIO4 CH04 | M12-2 pin 2 | Buffer conveyor sensor 2
    BUFFER_L4_STOPPER_RELAY_53RR7 AT %Q* : BOOL; // 48RIO4 CH05 | M12-3 pin 4 | 53RR7 coil, stopper motor #7 53M7, sheet 53.3/5A
    _48RIO4_SPARE_CH06 AT %Q* : BOOL; // 48RIO4 CH06 | M12-3 pin 2 | Spare
    BUFFER_L4_STOPPER_RELAY_53RR8 AT %Q* : BOOL; // 48RIO4 CH07 | M12-4 pin 4 | 53RR8 coil, sheet 53.3/7E (relay not detailed in drawing rev D)
    _48RIO4_SPARE_CH08 AT %Q* : BOOL; // 48RIO4 CH08 | M12-4 pin 2 | Spare
    _48RIO4_WcState AT %I* : BOOL; // DIO-05 > WcState > WcState (TRUE = data invalid)
    _48RIO4_EcState AT %I* : UINT; // DIO-05 > InfoData > State (8 = OP)

    // DIO-06 (EPP2328-0002) = 48RIO5 - conveyor with stopper, level 5 - sheets 48.5 and 53.4.
    BUFFER_L5_SAFETY_STOPPER_UPPER_SENSOR AT %I* : BOOL; // 48RIO5 CH01 | M12-1 pin 4 | Safety stopper upper sensor
    BUFFER_L5_SAFETY_STOPPER_LOWER_SENSOR AT %I* : BOOL; // 48RIO5 CH02 | M12-1 pin 2 | Safety stopper lower sensor
    BUFFER_L5_CONVEYOR_SENSOR_1 AT %I* : BOOL; // 48RIO5 CH03 | M12-2 pin 4 | Buffer conveyor sensor 1
    BUFFER_L5_CONVEYOR_SENSOR_2 AT %I* : BOOL; // 48RIO5 CH04 | M12-2 pin 2 | Buffer conveyor sensor 2
    BUFFER_L5_STOPPER_RELAY_53RR9 AT %Q* : BOOL; // 48RIO5 CH05 | M12-3 pin 4 | 53RR9 coil, stopper motor #9 53M9, sheet 53.4/5A
    _48RIO5_SPARE_CH06 AT %Q* : BOOL; // 48RIO5 CH06 | M12-3 pin 2 | Spare
    BUFFER_L5_STOPPER_RELAY_53RR10 AT %Q* : BOOL; // 48RIO5 CH07 | M12-4 pin 4 | 53RR10 coil, sheet 53.4/7E (relay not detailed in drawing rev D)
    _48RIO5_SPARE_CH08 AT %Q* : BOOL; // 48RIO5 CH08 | M12-4 pin 2 | Spare
    _48RIO5_WcState AT %I* : BOOL; // DIO-06 > WcState > WcState (TRUE = data invalid)
    _48RIO5_EcState AT %I* : UINT; // DIO-06 > InfoData > State (8 = OP)

    // DIO-07 (EPP2328-0002) = 48RIO6 - conveyor with stopper, level 6 - sheets 48.6 and 53.5.
    BUFFER_L6_SAFETY_STOPPER_UPPER_SENSOR AT %I* : BOOL; // 48RIO6 CH01 | M12-1 pin 4 | Safety stopper upper sensor
    BUFFER_L6_SAFETY_STOPPER_LOWER_SENSOR AT %I* : BOOL; // 48RIO6 CH02 | M12-1 pin 2 | Safety stopper lower sensor
    BUFFER_L6_CONVEYOR_SENSOR_1 AT %I* : BOOL; // 48RIO6 CH03 | M12-2 pin 4 | Buffer conveyor sensor 1
    BUFFER_L6_CONVEYOR_SENSOR_2 AT %I* : BOOL; // 48RIO6 CH04 | M12-2 pin 2 | Buffer conveyor sensor 2
    BUFFER_L6_STOPPER_RELAY_53RR11 AT %Q* : BOOL; // 48RIO6 CH05 | M12-3 pin 4 | 53RR11 coil, stopper motor #11 53M11, sheet 53.5/5A
    _48RIO6_SPARE_CH06 AT %Q* : BOOL; // 48RIO6 CH06 | M12-3 pin 2 | Spare
    BUFFER_L6_STOPPER_RELAY_53RR12 AT %Q* : BOOL; // 48RIO6 CH07 | M12-4 pin 4 | 53RR12 coil, sheet 53.5/7E (relay not detailed in drawing rev D)
    _48RIO6_SPARE_CH08 AT %Q* : BOOL; // 48RIO6 CH08 | M12-4 pin 2 | Spare
    _48RIO6_WcState AT %I* : BOOL; // DIO-07 > WcState > WcState (TRUE = data invalid)
    _48RIO6_EcState AT %I* : UINT; // DIO-07 > InfoData > State (8 = OP)

    // ---------------------------------------------------------------- TwinSAFE boxes
    // Safe channels travel in the FSoE frame to the TwinSAFE logic. They are NOT standard PLC I/O:
    // the standard PLC gets their state only through TwinSAFE logic outputs (IO_Safety).
    // Only diagnostics and the EP1957 standard (non-safe) data are declared here.

    // FDI-01 (EP1918-0002) = 43SRIO1 - safe inputs - sheets 43.0-43.1.
    //   In1/In2: 43SC1 to overtravel upper (NC).
    //   In3/In4: 43SC2 to overtravel lower (NC).
    //   In5-In8: spare.
    _43SRIO1_WcState AT %I* : BOOL; // FDI-01 > WcState > WcState (TRUE = data invalid)
    _43SRIO1_EcState AT %I* : UINT; // FDI-01 > InfoData > State (8 = OP)

    // FDIO-01 (EP1957-0022) = 43SRIO2 - safe inputs / outputs - sheets 43.2-43.4.
    //   In1/In2: 43LC1 light curtain receiver OSSD1 / OSSD2 (SICK C4C-EV13530B10000), sheet 43.4.
    //   In3/In4: 43LC2 light curtain sender (SICK C4C-SV13530B10000), sheet 43.4.
    //   Other safe inputs and safe outputs 1-4: not used in drawing rev D.
    _43SRIO2_SPARE_STD_OUT1 AT %Q* : BOOL; // FDIO-01 > Outputs > Module 1.Standard Output | Spare (no output used in drawing rev D)
    _43SRIO2_SPARE_STD_OUT2 AT %Q* : BOOL; // FDIO-01 > Outputs > Module 2.Standard Output | Spare (no output used in drawing rev D)
    _43SRIO2_SPARE_STD_OUT3 AT %Q* : BOOL; // FDIO-01 > Outputs > Module 3.Standard Output | Spare (no output used in drawing rev D)
    _43SRIO2_SPARE_STD_OUT4 AT %Q* : BOOL; // FDIO-01 > Outputs > Module 4.Standard Output | Spare (no output used in drawing rev D)
    _43SRIO2_FIELDVOLTAGE_UNDERRANGE AT %I* : BOOL; // FDIO-01 > FIELDVOLTAGE Field Voltage Status > Fieldvoltage Underrange
    _43SRIO2_FIELDVOLTAGE_OVERRANGE AT %I* : BOOL; // FDIO-01 > FIELDVOLTAGE Field Voltage Status > Fieldvoltage Overrange
    _43SRIO2_WcState AT %I* : BOOL; // FDIO-01 > WcState > WcState (TRUE = data invalid)
    _43SRIO2_EcState AT %I* : UINT; // FDIO-01 > InfoData > State (8 = OP)
END_VAR

// ---- GVLs/IO/IO_Safety.TcGVL
//{attribute 'qualified_only'}
VAR_GLOBAL
	ErrorAcknowledgement AT %Q*: BOOL;
	Run AT %Q*: BOOL;
END_VAR

// ---- GVLs/IO/IO_VFDs.TcGVL
{attribute 'qualified_only'}
VAR_GLOBAL
	
//---------------------------------------------------------VFD
    // VTD (MOVI-C MOVIPRO) / Module 1 (Standard 8 PD), MOVIKIT Positioning Drive.
    // Raw 16-bit UINT data, as defined in SpaceX.tsproj; no scaling or decoding.
    // Link each variable to the channel with the same number in TwinCAT XAE.
    // Word meanings from MOVISUITE; bit meanings and units still pending SEW.

    // Drive -> PLC: Inputs 8 PD / PDO 16#1A02 / object 16#7002.
    // Read only by FC Inputs, into Control.VTD.Motor.stProcessInput.
    VTD_PI_01 AT %I* : UINT; // PI 1, 16#7002:01 - Status word
    VTD_PI_02 AT %I* : UINT; // PI 2, 16#7002:02 - Actual speed
    VTD_PI_03 AT %I* : UINT; // PI 3, 16#7002:03 - Status/main fault - subfault
    VTD_PI_04 AT %I* : UINT; // PI 4, 16#7002:04 - Torque
    VTD_PI_05 AT %I* : UINT; // PI 5, 16#7002:05 - Digital inputs
    VTD_PI_06 AT %I* : UINT; // PI 6, 16#7002:06 - Actual application mode
    VTD_PI_07 AT %I* : UINT; // PI 7, 16#7002:07 - Actual position high word (DL50)
    VTD_PI_08 AT %I* : UINT; // PI 8, 16#7002:08 - Actual position low word (DL50)

    // PLC -> drive: Outputs 8 PD / PDO 16#1602 / object 16#6002.
    // Written only by FC Outputs, from Control.VTD.Motor.aProcessOutput.
    VTD_PO_01 AT %Q* : UINT; // PO 1, 16#6002:01 - Control word
    VTD_PO_02 AT %Q* : UINT; // PO 2, 16#6002:02 - Setpoint speed
    VTD_PO_03 AT %Q* : UINT; // PO 3, 16#6002:03 - Setpoint acceleration
    VTD_PO_04 AT %Q* : UINT; // PO 4, 16#6002:04 - Setpoint deceleration
    VTD_PO_05 AT %Q* : UINT; // PO 5, 16#6002:05 - Digital outputs
    VTD_PO_06 AT %Q* : UINT; // PO 6, 16#6002:06 - Setpoint application mode
    VTD_PO_07 AT %Q* : UINT; // PO 7, 16#6002:07 - Target position high word
    VTD_PO_08 AT %Q* : UINT; // PO 8, 16#6002:08 - Target position low word

    // EtherCAT diagnostics of the VTD box. Not linked yet: link manually in XAE.
    // Read only by FC Inputs.
    VTD_WcState AT %I* : BOOL; // VTD > WcState > WcState (TRUE = data invalid)
    VTD_EcState AT %I* : UINT; // VTD > InfoData > State (8 = OP)
	
	//----------------------------------------------------EXTRACTOR CONVEYOR
END_VAR
